// TIA Portal V21 export
VAR_GLOBAL   // PLC tag table "Default tag table"
   Start_Povoleno AT %I0.0 : Bool;
   Emergency_Stop AT %I0.1 : Bool;
   Ack AT %I0.2 : Bool;
   Fuse_OK AT %I0.3 : Bool;
   Horn AT %Q0.0 : Bool;
   Fault_Belt1 AT %M10.0 : Bool;
END_VAR
